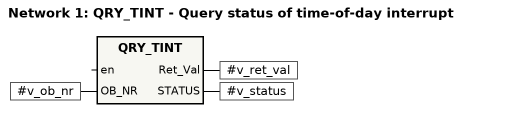
   #v_ret_val := QRY_TINT(OB_NR := #v_ob_nr, STATUS => #v_status);
END_REGION
END_FUNCTION_BLOCK

FUNCTION_BLOCK "FB_Fbd_ex109"   // FB121, FBD
{ S7_Optimized_Access := 'TRUE' }
   VAR_INPUT
      v_ob_nr : Int;
      v_dtime : Time;
      v_sign : Word;
   END_VAR
   VAR_OUTPUT
      v_ret_val : Int;
   END_VAR
BEGIN

REGION Network 1: SRT_DINT - Start time-delay interrupt
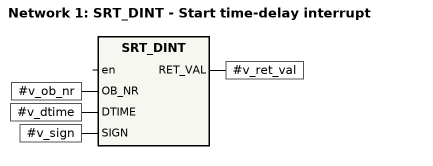
   #v_ret_val := SRT_DINT(OB_NR := #v_ob_nr, DTIME := #v_dtime, SIGN := #v_sign);
END_REGION
END_FUNCTION_BLOCK

FUNCTION_BLOCK "FB_Fbd_ex110"   // FB122, FBD
{ S7_Optimized_Access := 'TRUE' }
   VAR_INPUT
      v_ob_nr : Int;
   END_VAR
   VAR_OUTPUT
      v_ret_val : Int;
   END_VAR
BEGIN

REGION Network 1: CAN_DINT - Cancel time-delay interrupt
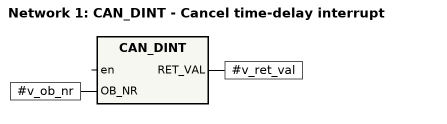
   #v_ret_val := CAN_DINT(OB_NR := #v_ob_nr);
END_REGION
END_FUNCTION_BLOCK

FUNCTION_BLOCK "FB_Fbd_ex111"   // FB123, FBD
{ S7_Optimized_Access := 'TRUE' }
   VAR_INPUT
      v_ob_nr : Int;
   END_VAR
   VAR_OUTPUT
      v_ret_val : Int;
      v_status : Word;
   END_VAR
BEGIN

REGION Network 1: QRY_DINT - Query time-delay interrupt status
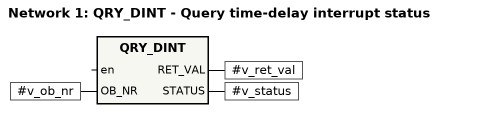
   #v_ret_val := QRY_DINT(OB_NR := #v_ob_nr, STATUS => #v_status);
END_REGION
END_FUNCTION_BLOCK

FUNCTION_BLOCK "FB_Fbd_ex112"   // FB124, FBD
{ S7_Optimized_Access := 'TRUE' }
   VAR_INPUT
      v_prgflt_set_mask : DWord;
      v_accflt_set_mask : DWord;
   END_VAR
   VAR_OUTPUT
      v_ret_val : Int;
      v_prgflt_masked : DWord;
      v_accflt_masked : DWord;
   END_VAR
BEGIN

REGION Network 1: MSK_FLT - Mask synchronous error events
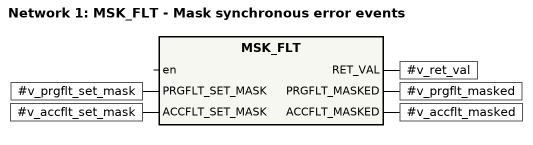
   #v_ret_val := MSK_FLT(PRGFLT_SET_MASK := #v_prgflt_set_mask,
                         ACCFLT_SET_MASK := #v_accflt_set_mask,
                         PRGFLT_MASKED => #v_prgflt_masked,
                         ACCFLT_MASKED => #v_accflt_masked);
END_REGION
END_FUNCTION_BLOCK

FUNCTION_BLOCK "FB_Fbd_ex113"   // FB125, FBD
{ S7_Optimized_Access := 'TRUE' }
   VAR_INPUT
      v_prgflt_reset_mask : DWord;
      v_accflt_reset_mask : DWord;
   END_VAR
   VAR_OUTPUT
      v_ret_val : Int;
      v_prgflt_masked : DWord;
      v_accflt_masked : DWord;
   END_VAR
BEGIN

REGION Network 1: DMSK_FLT - Unmask synchronous error events
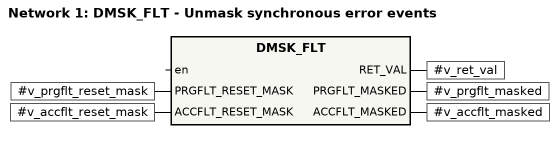
   #v_ret_val := DMSK_FLT(PRGFLT_RESET_MASK := #v_prgflt_reset_mask,
                          ACCFLT_RESET_MASK := #v_accflt_reset_mask,
                          PRGFLT_MASKED => #v_prgflt_masked,
                          ACCFLT_MASKED => #v_accflt_masked);
END_REGION
END_FUNCTION_BLOCK

FUNCTION_BLOCK "FB_Fbd_ex114"   // FB126, FBD
{ S7_Optimized_Access := 'TRUE' }
   VAR_INPUT
      v_prgflt_query : DWord;
      v_accflt_query : DWord;
   END_VAR
   VAR_OUTPUT
      v_ret_val : Int;
      v_prgflt_clr : DWord;
      v_accflt_clr : DWord;
   END_VAR
BEGIN

REGION Network 1: READ_ERR - Read out event status register
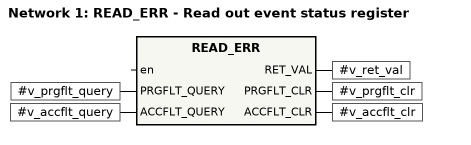
   #v_ret_val := READ_ERR(PRGFLT_QUERY := #v_prgflt_query,
                          ACCFLT_QUERY := #v_accflt_query,
                          PRGFLT_CLR => #v_prgflt_clr,
                          ACCFLT_CLR => #v_accflt_clr);
END_REGION
END_FUNCTION_BLOCK

FUNCTION_BLOCK "FB_Fbd_ex115"   // FB127, FBD
{ S7_Optimized_Access := 'TRUE' }
   VAR_INPUT
      v_mode : Byte;
      v_ob_nr : Int;
   END_VAR
   VAR_OUTPUT
      v_ret_val : Int;
   END_VAR
BEGIN

REGION Network 1: DIS_IRT - Disable interrupt event
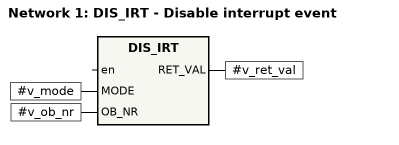
   #v_ret_val := DIS_IRT(MODE := #v_mode, OB_NR := #v_ob_nr);
END_REGION
END_FUNCTION_BLOCK

FUNCTION_BLOCK "FB_Fbd_ex116"   // FB128, FBD
{ S7_Optimized_Access := 'TRUE' }
   VAR_INPUT
      v_mode : Byte;
      v_ob_nr : Int;
   END_VAR
   VAR_OUTPUT
      v_ret_val : Int;
   END_VAR
BEGIN

REGION Network 1: EN_IRT - Enable interrupt event
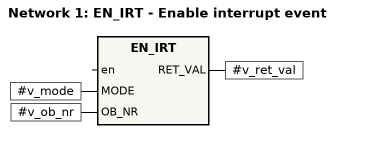
   #v_ret_val := EN_IRT(MODE := #v_mode, OB_NR := #v_ob_nr);
END_REGION
END_FUNCTION_BLOCK

FUNCTION_BLOCK "FB_Fbd_ex117"   // FB129, FBD
{ S7_Optimized_Access := 'TRUE' }
   VAR_OUTPUT
      v_ret_val : Int;
   END_VAR
BEGIN

REGION Network 1: DIS_AIRT - Delay execution of higher priority interrupts and asynchronous error events
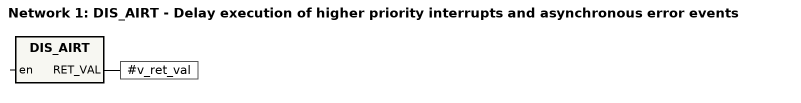
   #v_ret_val := DIS_AIRT();
END_REGION
END_FUNCTION_BLOCK

FUNCTION_BLOCK "FB_Fbd_ex118"   // FB130, FBD
{ S7_Optimized_Access := 'TRUE' }
   VAR_OUTPUT
      v_ret_val : Int;
   END_VAR
BEGIN

REGION Network 1: EN_AIRT - Enable execution of higher priority interrupts and asynchronous error events
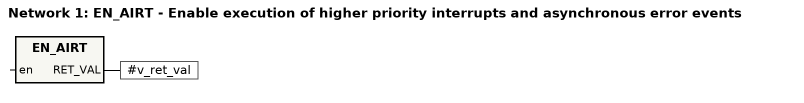
   #v_ret_val := EN_AIRT();
END_REGION
END_FUNCTION_BLOCK

FUNCTION_BLOCK "FB_Fbd_ex120"   // FB131, FBD
{ S7_Optimized_Access := 'TRUE' }
   VAR_INPUT
      v_alarm : ALARM_BASE;
   END_VAR
   VAR_OUTPUT
      v_alarmstate : Byte;
      v_error : Bool;
      v_status : Word;
   END_VAR
BEGIN

REGION Network 1: Get_AlarmState - Output alarm status
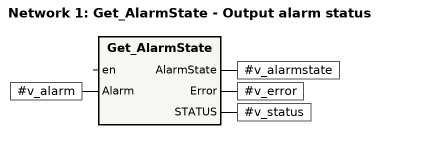
   // no SCL statement known for Get_AlarmState: written as a call
   Get_AlarmState(Alarm := #v_alarm, AlarmState => #v_alarmstate, Error => #v_error, STATUS => #v_status);
END_REGION
END_FUNCTION_BLOCK

FUNCTION_BLOCK "FB_Fbd_ex121"   // FB132, FBD
{ S7_Optimized_Access := 'TRUE' }
   VAR_INPUT
      v_mode : UInt;
      v_textid : UInt;
      v_textlistid : UInt;
   END_VAR
   VAR_OUTPUT
      v_ret_val : Int;
   END_VAR
   VAR_IN_OUT
      v_assocvalues : AssocValues;
   END_VAR
BEGIN

REGION Network 1: Gen_UsrMsg - Generate user diagnostic alarms
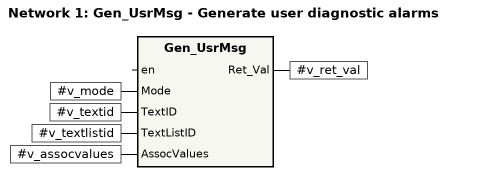
   // no SCL statement known for Gen_UsrMsg: written as a call
   #v_ret_val := Gen_UsrMsg(Mode := #v_mode,
                           TextID := #v_textid,
                           TextListID := #v_textlistid,
                           AssocValues := #v_assocvalues);
END_REGION
END_FUNCTION_BLOCK

FUNCTION_BLOCK "FB_Fbd_ex123"   // FB133, FBD
{ S7_Optimized_Access := 'TRUE' }
   VAR_INPUT
      v_mode : UInt;
   END_VAR
   VAR_OUTPUT
      v_error : Bool;
      v_status : Word;
   END_VAR
BEGIN

REGION Network 1: Ack_Alarms - Acknowledge alarms
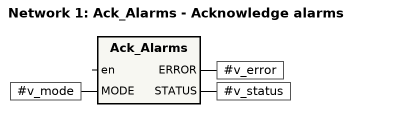
   // no SCL statement known for Ack_Alarms: written as a call
   Ack_Alarms(MODE := #v_mode, ERROR => #v_error, STATUS => #v_status);
END_REGION
END_FUNCTION_BLOCK

FUNCTION_BLOCK "FB_Fbd_ex124"   // FB134, FBD
{ S7_Optimized_Access := 'TRUE' }
   VAR_OUTPUT
      v_ret_val : Int;
   END_VAR
   VAR_IN_OUT
      v_top_si : Array[0..99] of Byte;
      v_start_up_si : Array[0..99] of Byte;
   END_VAR
BEGIN

REGION Network 1: RD_SINFO - Read current OB start information
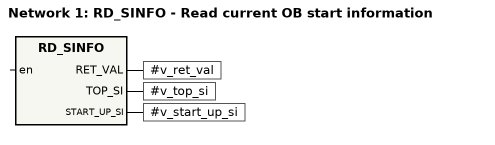
   #v_ret_val := RD_SINFO(TOP_SI => #v_top_si, START_UP_SI => #v_start_up_si);
END_REGION
END_FUNCTION_BLOCK

FUNCTION_BLOCK "FB_Fbd_ex125"   // FB135, FBD
{ S7_Optimized_Access := 'TRUE' }
   VAR_INPUT
      v_mode : UInt;
      v_ob : OB_Any;
   END_VAR
   VAR_OUTPUT
      v_ret_val : Int;
   END_VAR
   VAR_IN_OUT
      v_info : Variant;
   END_VAR
BEGIN

REGION Network 1: RT_INFO - Read out runtime statistics
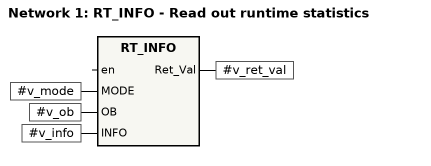
   #v_ret_val := RT_INFO(MODE := #v_mode, OB := #v_ob, INFO := #v_info);
END_REGION
END_FUNCTION_BLOCK

FUNCTION_BLOCK "FB_Fbd_ex126"   // FB136, FBD
{ S7_Optimized_Access := 'TRUE' }
   VAR_INPUT
      v_laddr : Hw_Io;
      v_led : UInt;
   END_VAR
   VAR_OUTPUT
      v_ret_val : Int;
   END_VAR
BEGIN

REGION Network 1: LED - Read LED status
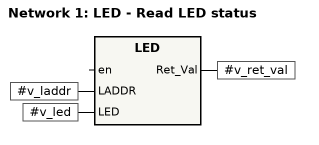
   #v_ret_val := LED(LADDR := #v_laddr, LED := #v_led);
END_REGION
END_FUNCTION_BLOCK

FUNCTION_BLOCK "FB_Fbd_ex127"   // FB137, FBD
{ S7_Optimized_Access := 'TRUE' }
   VAR_INPUT
      v_laddr : Hw_Io;
      v_im_type : UInt;
   END_VAR
   VAR_OUTPUT
      v_done : Bool;
      v_busy : Bool;
      v_error : Bool;
      v_status : Word;
   END_VAR
   VAR_IN_OUT
      v_data : Array[0..99] of Byte;
   END_VAR
   VAR
      inst : Get_IM_Data;
   END_VAR
BEGIN

REGION Network 1: Get_IM_Data - Reading identification and maintenance data
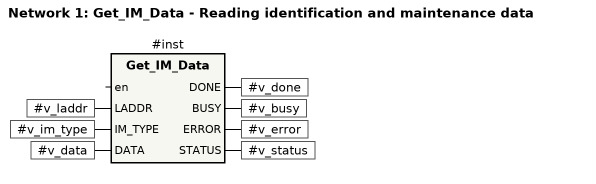
   #inst(LADDR := #v_laddr,   // Get_IM_Data
         IM_TYPE := #v_im_type,
         DATA := #v_data,
         DONE => #v_done,
         BUSY => #v_busy,
         ERROR => #v_error,
         STATUS => #v_status);
END_REGION
END_FUNCTION_BLOCK

FUNCTION_BLOCK "FB_Fbd_ex128"   // FB138, FBD
{ S7_Optimized_Access := 'TRUE' }
   VAR_INPUT
      v_laddr : Hw_IoSystem;
      v_station_nr : UInt;
   END_VAR
   VAR_OUTPUT
      v_done : Bool;
      v_busy : Bool;
      v_error : Bool;
      v_len : DInt;
      v_status : Word;
   END_VAR
   VAR_IN_OUT
      v_data : Array[0..99] of Byte;
   END_VAR
   VAR
      inst : Get_Name;
   END_VAR
BEGIN

REGION Network 1: GET_NAME - Read out name of an IO device or a DP slave
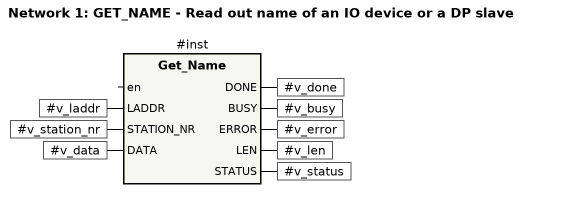
   #inst(LADDR := #v_laddr,   // Get_Name
         STATION_NR := #v_station_nr,
         DATA := #v_data,
         DONE => #v_done,
         BUSY => #v_busy,
         ERROR => #v_error,
         LEN => #v_len,
         STATUS => #v_status);
END_REGION
END_FUNCTION_BLOCK

FUNCTION_BLOCK "FB_Fbd_ex129"   // FB139, FBD
{ S7_Optimized_Access := 'TRUE' }
   VAR_INPUT
      v_req : Bool;
      v_laddr : Hw_Device;
      v_detail : Hw_SubModule;
      v_mode : UInt;
   END_VAR
   VAR_OUTPUT
      v_done : Bool;
      v_busy : Bool;
      v_error : Bool;
      v_status : Word;
   END_VAR
   VAR_IN_OUT
      v_data : Array[0..99] of Byte;
   END_VAR
   VAR
      inst : GetStationInfo;
   END_VAR
BEGIN

REGION Network 1: GetStationInfo - Read information of an IO device
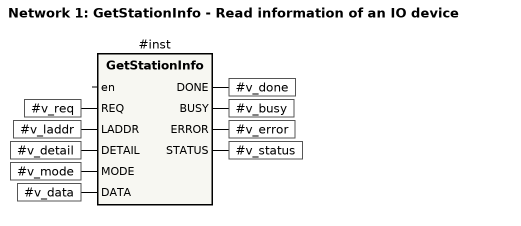
   #inst(REQ := #v_req,   // GetStationInfo
         LADDR := #v_laddr,
         DETAIL := #v_detail,
         MODE := #v_mode,
         DATA := #v_data,
         DONE => #v_done,
         BUSY => #v_busy,
         ERROR => #v_error,
         STATUS => #v_status);
END_REGION
END_FUNCTION_BLOCK

FUNCTION_BLOCK "FB_Fbd_ex130"   // FB140, FBD
{ S7_Optimized_Access := 'TRUE' }
   VAR_INPUT
      v_laddr : Hw_IoSystem;
      v_mode : UInt;
   END_VAR
   VAR_OUTPUT
      v_ret_val : Int;
   END_VAR
   VAR_IN_OUT
      v_state : Variant;
   END_VAR
BEGIN

REGION Network 1: DeviceStates - Read module status information in an IO system
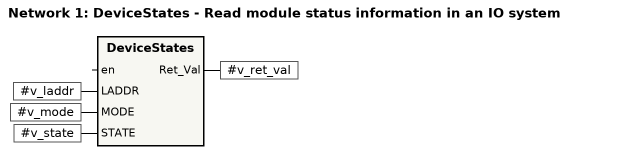
   // no SCL statement known for DeviceStates: written as a call
   #v_ret_val := DeviceStates(LADDR := #v_laddr, MODE := #v_mode, STATE := #v_state);
END_REGION
END_FUNCTION_BLOCK

FUNCTION_BLOCK "FB_Fbd_ex131"   // FB141, FBD
{ S7_Optimized_Access := 'TRUE' }
   VAR_INPUT
      v_laddr : Hw_Device;
      v_mode : UInt;
   END_VAR
   VAR_OUTPUT
      v_ret_val : Int;
   END_VAR
   VAR_IN_OUT
      v_state : Variant;
   END_VAR
BEGIN

REGION Network 1: ModuleStates - Read module status information of a module
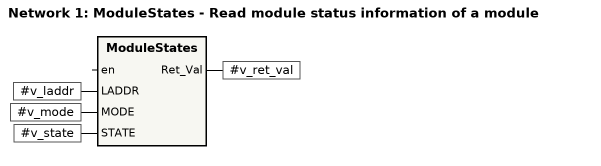
   // no SCL statement known for ModuleStates: written as a call
   #v_ret_val := ModuleStates(LADDR := #v_laddr, MODE := #v_mode, STATE := #v_state);
END_REGION
END_FUNCTION_BLOCK

FUNCTION_BLOCK "FB_Fbd_ex132"   // FB142, FBD
{ S7_Optimized_Access := 'TRUE' }
   VAR_INPUT
      v_laddr : Hw_Any;
      v_mode : UInt;
   END_VAR
   VAR_OUTPUT
      v_ret_val : Int;
   END_VAR
   VAR_IN_OUT
      v_diagevent : DiagnosticDetail;
   END_VAR
BEGIN

REGION Network 1: GEN_DIAG - Generate diagnostics information
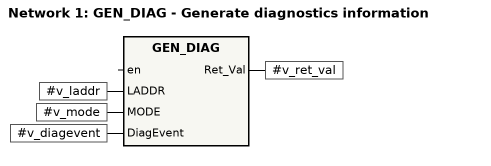
   #v_ret_val := GEN_DIAG(LADDR := #v_laddr, MODE := #v_mode, DiagEvent := #v_diagevent);
END_REGION
END_FUNCTION_BLOCK

FUNCTION_BLOCK "FB_Fbd_ex133"   // FB143, FBD
{ S7_Optimized_Access := 'TRUE' }
   VAR_INPUT
      v_mode : UInt;
      v_laddr : Hw_Any;
   END_VAR
   VAR_OUTPUT
      v_ret_val : Int;
      v_cnt_diag : UInt;
   END_VAR
   VAR_IN_OUT
      v_diag : Variant;
      v_detail : Variant;
   END_VAR
BEGIN

REGION Network 1: GET_DIAG - Read diagnostic information
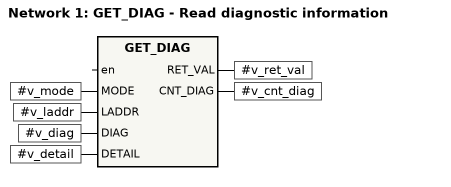
   #v_ret_val := GET_DIAG(MODE := #v_mode,
                          LADDR := #v_laddr,
                          DIAG := #v_diag,
                          DETAIL := #v_detail,
                          CNT_DIAG => #v_cnt_diag);
END_REGION
END_FUNCTION_BLOCK

FUNCTION_BLOCK "FB_Fbd_ex135"   // FB144, FBD
{ S7_Optimized_Access := 'TRUE' }
   VAR_INPUT
      v_req : Bool;
   END_VAR
   VAR_OUTPUT
      v_done : Bool;
      v_busy : Bool;
      v_error : Bool;
      v_status : Word;
   END_VAR
   VAR_IN_OUT
      v_recipe_db : Array[0..99] of Byte;
   END_VAR
   VAR
      inst : RecipeExport;
   END_VAR
BEGIN

REGION Network 1: RecipeExport - Exporting recipes
